Fanuc KAREL source: kt00573.KL

-- PROVISIONAL review KL for V770-1; original PC SHA256 c10f4c959a81e2d7cb84ae5d6c3d74fe73aab11ce54f3449cfbf8c4edfb5b6e5
-- Incomplete behavior may be omitted. Consult companion uncertainty JSON. Do not deploy.
PROGRAM KT00573
%NOLOCKGROUP
VAR
  R1 : REAL
-- UNRESOLVED_DECL V2 type=000013
-- UNRESOLVED_DECL OUT type=000013
BEGIN
  -- UNRESOLVED_PC offsets 5-16; opcodes 2E,23
  -- UNRESOLVED_PC offsets 21-36; opcodes 2E,22,32,35
  -- UNRESOLVED_PC offsets 41-63; opcodes 21,49,8C,4A
  -- UNRESOLVED_PC offsets 68-72; opcodes 7F
END KT00573
